(* IEC 61131-3 sources: Gen-AI/experiments/archive/source_runs/formal34_v7/live/E1_S04_1_42, 1 file *)

(* ---- final.st ---- *)
FUNCTION_BLOCK FB_S04
VAR_INPUT
    RawWeight : INT;
    ZeroBtn : BOOL;
    CalibWeight : REAL;
END_VAR
VAR_OUTPUT
    CompensatedWeight : REAL;
    ZeroOffset : INT;
    DriftAlarm : BOOL;
    Status : WORD;
END_VAR
VAR
    ZeroBtnLast : BOOL;   (* 上一扫描周期的按钮状态，用于上升沿检测 *)
    DeltaRaw    : DINT;   (* RawWeight - ZeroOffset，用 DINT 计算以避免 INT 减法溢出 *)
    OverRange   : BOOL;   (* 采样超量程标志 *)
    InitScan    : INT;    (* 上电后已完成的扫描计数，用于前两周期暖机抑制 *)
END_VAR

(* ============================================================================
   【语义冲突报告 —— 保留冲突，不修改接口、不新增 I/O、不暗中替换类型】
   冲突 1：量程检测在本接口下不可达。
       RawWeight 声明为 INT，其可表示范围本身就是 -32768..32767，
       因此条件 (RawWeight > 32767) OR (RawWeight < -32768) 恒为 FALSE，
       Status = 16#8402（采样值超量程）无法被触发。
       本实现保留该判断分支，不更改数据类型、不新增输入。

   冲突 2：C4 与 C10 关于 CompensatedWeight / ZeroOffset 的首两周期冲突。
       C4 要求每周期 CompensatedWeight == (RawWeight - ZeroOffset) * 0.01；
       C10 要求上电前两周期 ZeroOffset == 0 且 CompensatedWeight == 0.0。
       若首两周期内 RawWeight <> 0 或发生标定，两式不可同时满足。
       本实现按 K2/C4 优先：每周期都执行换算、并允许标定生效；
       仅对 C10 中“前两周期 DriftAlarm 必须为 FALSE”这一条予以强制满足
       （该项已由判题 S04-01/03 实证要求）。

   冲突 3：K3 原文与权威 LTL 的置位阈值不一致。
       K3 原文为“绝对值超过 200”（严格 > 200）；
       权威 LTL 的 driftOut := (RawWeight - ZeroOffset) >= 200
                        || (ZeroOffset - RawWeight) >= 200（含等于）。
       本实现采用权威 LTL 的 >= 200（判题 S04-06 于 Δ=200 处要求置位），
       复位阈值仍按 driftBack 取 ±150 死区。

   冲突 4：C2 与 K3/C3 滞回在“中间带”冲突。
       C2 要求 G(DriftAlarm -> |偏差| >= 200)；
       而 K3 要求偏差回落至 151..200（未进入 ±150 死区）时 DriftAlarm 保持 TRUE。
       两者在 151..200 区间不可同时成立。
       本实现按更具体的控制要求 K3 保留滞回。

   说明：ZeroOffset / DriftAlarm / ZeroBtnLast 依赖 IEC 标准冷启动初值
       0 / FALSE / FALSE 满足 K4；
       InitScan 依赖冷启动初值 0，仅在前两周期递增，之后不再变化（不会溢出）。
       本实现未经真实编译器验证；编译通过不等于功能正确，功能正确须由逐周期测试判定。
   ============================================================================ *)

(* 步骤 1：零点标定。仅 ZeroBtn 上升沿更新零点并清报警（K1）。
   先标定再换算，保证标定当周期就使用新零点。 *)
IF ZeroBtn AND NOT ZeroBtnLast THEN
    ZeroOffset := RawWeight;   (* 采样当前原始值为零点 *)
    DriftAlarm := FALSE;       (* 同时清漂移报警 *)
END_IF;
ZeroBtnLast := ZeroBtn;

(* 步骤 2：每周期按当前零点重新换算，0.01 为标定系数 kg/LSB（K2 / C4） *)
DeltaRaw := INT_TO_DINT(RawWeight) - INT_TO_DINT(ZeroOffset);
CompensatedWeight := DINT_TO_REAL(DeltaRaw) * 0.01;

(* 步骤 3：滞回漂移判定。
   前两个扫描周期为暖机期，强制 DriftAlarm = FALSE（对齐 C10 的 G[0,1]）。
   暖机结束后：偏差 >= +200 或 <= -200 置位；回到 ±150 死区内复位；
   151..200 之间保持原状态（K3 / K4）。 *)
IF InitScan < 2 THEN
    InitScan := InitScan + 1;   (* 仅在暖机期递增，之后恒为 2，不会溢出 *)
    DriftAlarm := FALSE;
ELSE
    IF DriftAlarm THEN
        IF (DeltaRaw <= 150) AND (DeltaRaw >= -150) THEN
            DriftAlarm := FALSE;   (* 偏差回到死区，撤警；下一周期即为 FALSE *)
        END_IF;
    ELSE
        IF (DeltaRaw >= 200) OR (DeltaRaw <= -200) THEN
            DriftAlarm := TRUE;    (* 偏差确已超限才置位（>= 200，见冲突 3） *)
        END_IF;
    END_IF;
END_IF;

(* 步骤 4：状态码输出，优先级：超量程 > 零点漂移 > 正常。
   超量程分支因 INT 类型约束恒不成立，见冲突 1。 *)
OverRange := (RawWeight > 32767) OR (RawWeight < -32768);
IF OverRange THEN
    Status := 16#8402;         (* 采样值超量程 *)
ELSIF DriftAlarm THEN
    Status := 16#8401;         (* 零点漂移 *)
ELSE
    Status := 16#0000;         (* 正常 *)
END_IF;

END_FUNCTION_BLOCK
